(*
SPDX-FileCopyrightText: © 2026 Oleksandr Tiutyk <trofimich@gmail.com>
SPDX-License-Identifier: MIT
License: https://opensource.org/license/mit
*)

(*!
<summary>Describes the original IEC type and shape of one owned declaration.</summary>
<description>ElementSize includes the terminator and full capacity for STRING or WSTRING. ElementCount is always positive.
IsArray distinguishes a scalar from a single-element array.</description>
*)
TYPE VARIABLE_DECLARATION :
STRUCT
	ElementType : __SYSTEM.TYPE_CLASS;
	ElementSize : UDINT;
	ElementCount : DINT;
	IsArray : BOOL;
END_STRUCT
END_TYPE

(* stored: Version 1.1.0.1
   DUT VARIABLE_DECLARATION: Id {19111c89-5249-4cbb-8df5-91ef7f39f05a} *)
